// TIA Portal V19 export
FUNCTION_BLOCK "ALL_AI"   // FB2, FBD
{ S7_Optimized_Access := 'TRUE' }
// stored: MemoryReserve 100, SetENOAutomatically false
   VAR
      AI_TT01 { S7_SetPoint := 'True'} : "AI";
      TT_01 { S7_SetPoint := 'True'} : "AI";
      TT_02 { S7_SetPoint := 'True'} : "AI";
      TT_03 { S7_SetPoint := 'True'} : "AI";
      APT01 { S7_SetPoint := 'True'} : "AI";
      GPT01 { S7_SetPoint := 'True'} : "AI";
      GPT02 { S7_SetPoint := 'True'} : "AI";
      GPT03 { S7_SetPoint := 'True'} : "AI";
      GPT04 { S7_SetPoint := 'True'} : "AI";
      O201 { S7_SetPoint := 'True'} : "AI";
      LEL01 { S7_SetPoint := 'True'} : "AI";
      LEL02 { S7_SetPoint := 'True'} : "AI";
      PS01 { S7_SetPoint := 'True'} : "AI";
      RLT01 { S7_SetPoint := 'True'} : "AI";
      Weighing { S7_SetPoint := 'True'} : "AI";
   END_VAR
BEGIN

REGION Network 1: TT01
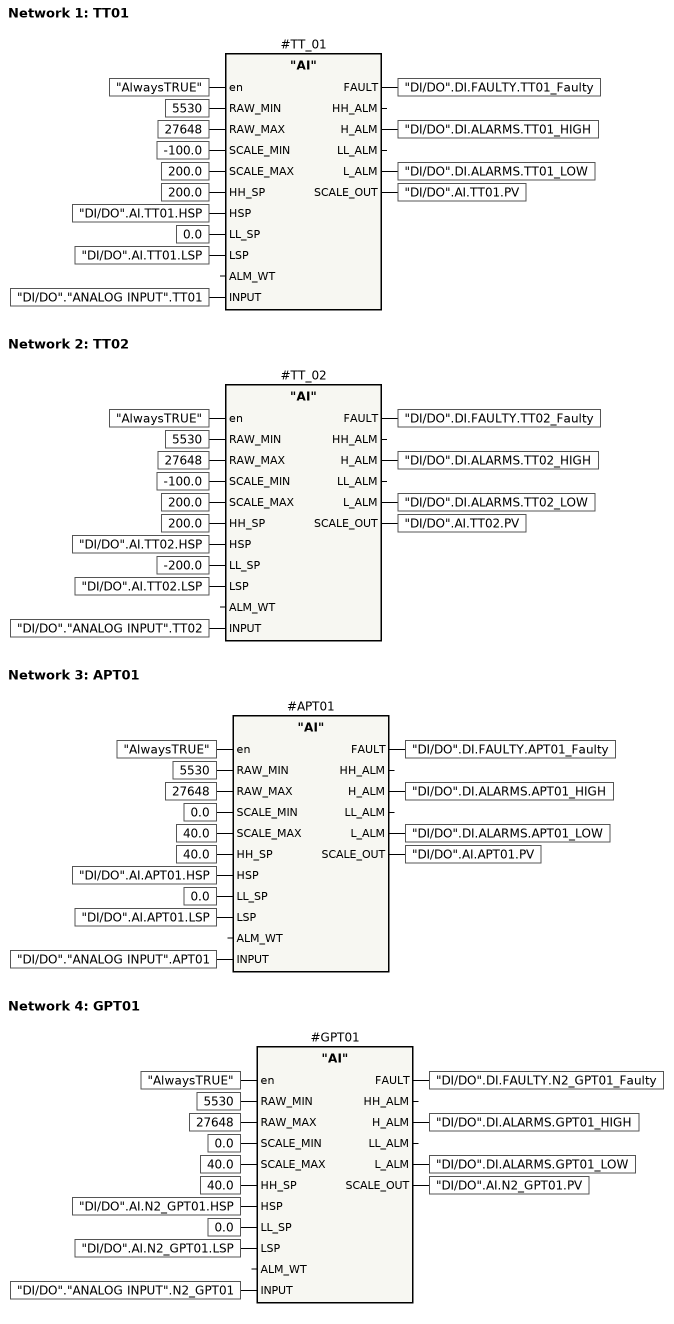
   IF "AlwaysTRUE" THEN
       #TT_01(RAW_MIN := 5530,   // "AI"
              RAW_MAX := 27648,
              SCALE_MIN := -100.0,
              SCALE_MAX := 200.0,
              HH_SP := 200.0,
              HSP := "DI/DO".AI.TT01.HSP,
              LL_SP := 0.0,
              LSP := "DI/DO".AI.TT01.LSP,
              INPUT := "DI/DO"."ANALOG INPUT".TT01,
              FAULT => "DI/DO".DI.FAULTY.TT01_Faulty,
              H_ALM => "DI/DO".DI.ALARMS.TT01_HIGH,
              L_ALM => "DI/DO".DI.ALARMS.TT01_LOW,
              SCALE_OUT => "DI/DO".AI.TT01.PV);
   END_IF;
END_REGION

REGION Network 2: TT02
   IF "AlwaysTRUE" THEN
       #TT_02(RAW_MIN := 5530,   // "AI"
              RAW_MAX := 27648,
              SCALE_MIN := -100.0,
              SCALE_MAX := 200.0,
              HH_SP := 200.0,
              HSP := "DI/DO".AI.TT02.HSP,
              LL_SP := -200.0,
              LSP := "DI/DO".AI.TT02.LSP,
              INPUT := "DI/DO"."ANALOG INPUT".TT02,
              FAULT => "DI/DO".DI.FAULTY.TT02_Faulty,
              H_ALM => "DI/DO".DI.ALARMS.TT02_HIGH,
              L_ALM => "DI/DO".DI.ALARMS.TT02_LOW,
              SCALE_OUT => "DI/DO".AI.TT02.PV);
   END_IF;
END_REGION

REGION Network 3: APT01
   IF "AlwaysTRUE" THEN
       #APT01(RAW_MIN := 5530,   // "AI"
              RAW_MAX := 27648,
              SCALE_MIN := 0.0,
              SCALE_MAX := 40.0,
              HH_SP := 40.0,
              HSP := "DI/DO".AI.APT01.HSP,
              LL_SP := 0.0,
              LSP := "DI/DO".AI.APT01.LSP,
              INPUT := "DI/DO"."ANALOG INPUT".APT01,
              FAULT => "DI/DO".DI.FAULTY.APT01_Faulty,
              H_ALM => "DI/DO".DI.ALARMS.APT01_HIGH,
              L_ALM => "DI/DO".DI.ALARMS.APT01_LOW,
              SCALE_OUT => "DI/DO".AI.APT01.PV);
   END_IF;
END_REGION

REGION Network 4: GPT01
   IF "AlwaysTRUE" THEN
       #GPT01(RAW_MIN := 5530,   // "AI"
              RAW_MAX := 27648,
              SCALE_MIN := 0.0,
              SCALE_MAX := 40.0,
              HH_SP := 40.0,
              HSP := "DI/DO".AI.N2_GPT01.HSP,
              LL_SP := 0.0,
              LSP := "DI/DO".AI.N2_GPT01.LSP,
              INPUT := "DI/DO"."ANALOG INPUT".N2_GPT01,
              FAULT => "DI/DO".DI.FAULTY.N2_GPT01_Faulty,
              H_ALM => "DI/DO".DI.ALARMS.GPT01_HIGH,
              L_ALM => "DI/DO".DI.ALARMS.GPT01_LOW,
              SCALE_OUT => "DI/DO".AI.N2_GPT01.PV);
   END_IF;
END_REGION

REGION Network 5: GPT02
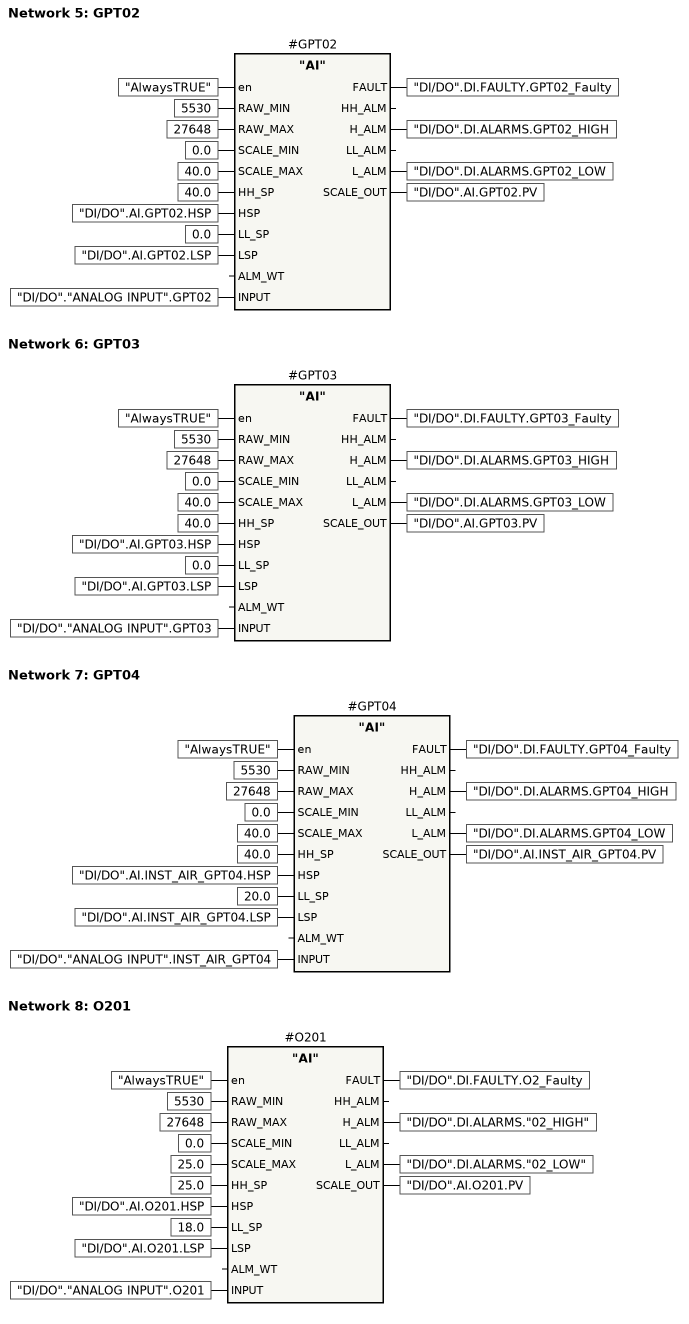
   IF "AlwaysTRUE" THEN
       #GPT02(RAW_MIN := 5530,   // "AI"
              RAW_MAX := 27648,
              SCALE_MIN := 0.0,
              SCALE_MAX := 40.0,
              HH_SP := 40.0,
              HSP := "DI/DO".AI.GPT02.HSP,
              LL_SP := 0.0,
              LSP := "DI/DO".AI.GPT02.LSP,
              INPUT := "DI/DO"."ANALOG INPUT".GPT02,
              FAULT => "DI/DO".DI.FAULTY.GPT02_Faulty,
              H_ALM => "DI/DO".DI.ALARMS.GPT02_HIGH,
              L_ALM => "DI/DO".DI.ALARMS.GPT02_LOW,
              SCALE_OUT => "DI/DO".AI.GPT02.PV);
   END_IF;
END_REGION

REGION Network 6: GPT03
   IF "AlwaysTRUE" THEN
       #GPT03(RAW_MIN := 5530,   // "AI"
              RAW_MAX := 27648,
              SCALE_MIN := 0.0,
              SCALE_MAX := 40.0,
              HH_SP := 40.0,
              HSP := "DI/DO".AI.GPT03.HSP,
              LL_SP := 0.0,
              LSP := "DI/DO".AI.GPT03.LSP,
              INPUT := "DI/DO"."ANALOG INPUT".GPT03,
              FAULT => "DI/DO".DI.FAULTY.GPT03_Faulty,
              H_ALM => "DI/DO".DI.ALARMS.GPT03_HIGH,
              L_ALM => "DI/DO".DI.ALARMS.GPT03_LOW,
              SCALE_OUT => "DI/DO".AI.GPT03.PV);
   END_IF;
END_REGION

REGION Network 7: GPT04
   IF "AlwaysTRUE" THEN
       #GPT04(RAW_MIN := 5530,   // "AI"
              RAW_MAX := 27648,
              SCALE_MIN := 0.0,
              SCALE_MAX := 40.0,
              HH_SP := 40.0,
              HSP := "DI/DO".AI.INST_AIR_GPT04.HSP,
              LL_SP := 20.0,
              LSP := "DI/DO".AI.INST_AIR_GPT04.LSP,
              INPUT := "DI/DO"."ANALOG INPUT".INST_AIR_GPT04,
              FAULT => "DI/DO".DI.FAULTY.GPT04_Faulty,
              H_ALM => "DI/DO".DI.ALARMS.GPT04_HIGH,
              L_ALM => "DI/DO".DI.ALARMS.GPT04_LOW,
              SCALE_OUT => "DI/DO".AI.INST_AIR_GPT04.PV);
   END_IF;
END_REGION

REGION Network 8: O201
   IF "AlwaysTRUE" THEN
       #O201(RAW_MIN := 5530,   // "AI"
             RAW_MAX := 27648,
             SCALE_MIN := 0.0,
             SCALE_MAX := 25.0,
             HH_SP := 25.0,
             HSP := "DI/DO".AI.O201.HSP,
             LL_SP := 18.0,
             LSP := "DI/DO".AI.O201.LSP,
             INPUT := "DI/DO"."ANALOG INPUT".O201,
             FAULT => "DI/DO".DI.FAULTY.O2_Faulty,
             H_ALM => "DI/DO".DI.ALARMS."02_HIGH",
             L_ALM => "DI/DO".DI.ALARMS."02_LOW",
             SCALE_OUT => "DI/DO".AI.O201.PV);
   END_IF;
END_REGION

REGION Network 9: LEL01
   // Configuration pending
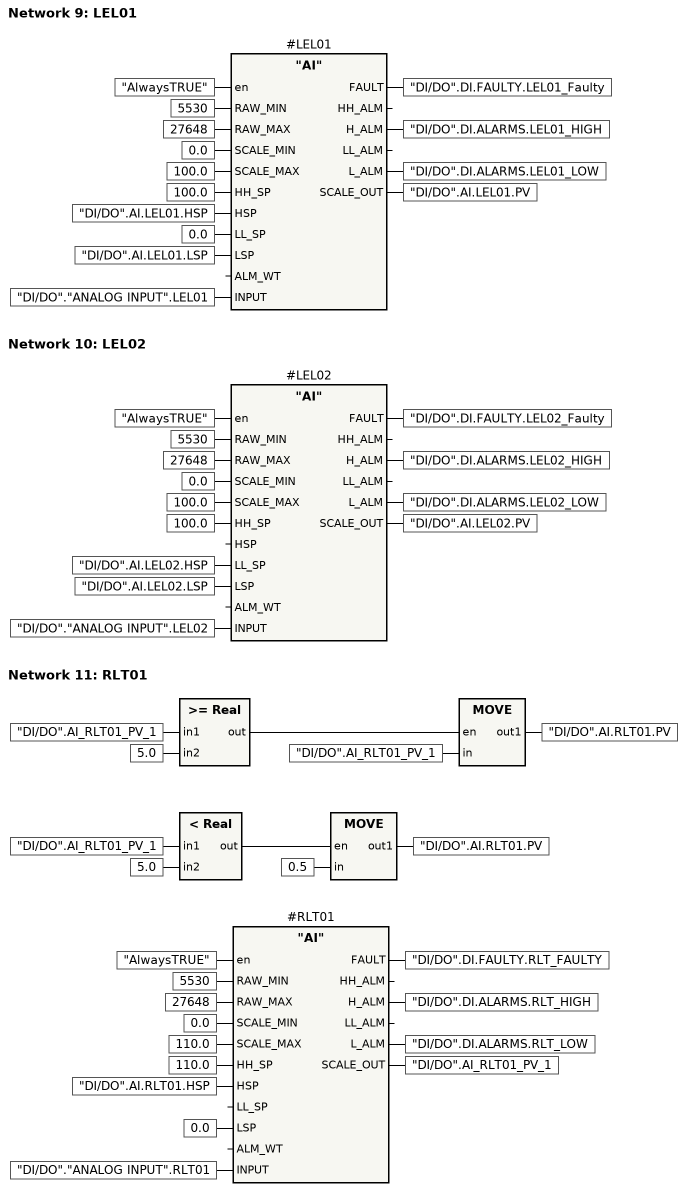
   IF "AlwaysTRUE" THEN
       #LEL01(RAW_MIN := 5530,   // "AI"
              RAW_MAX := 27648,
              SCALE_MIN := 0.0,
              SCALE_MAX := 100.0,
              HH_SP := 100.0,
              HSP := "DI/DO".AI.LEL01.HSP,
              LL_SP := 0.0,
              LSP := "DI/DO".AI.LEL01.LSP,
              INPUT := "DI/DO"."ANALOG INPUT".LEL01,
              FAULT => "DI/DO".DI.FAULTY.LEL01_Faulty,
              H_ALM => "DI/DO".DI.ALARMS.LEL01_HIGH,
              L_ALM => "DI/DO".DI.ALARMS.LEL01_LOW,
              SCALE_OUT => "DI/DO".AI.LEL01.PV);
   END_IF;
END_REGION

REGION Network 10: LEL02
   // Instrument is not installed at site
   IF "AlwaysTRUE" THEN
       #LEL02(RAW_MIN := 5530,   // "AI"
              RAW_MAX := 27648,
              SCALE_MIN := 0.0,
              SCALE_MAX := 100.0,
              HH_SP := 100.0,
              LL_SP := "DI/DO".AI.LEL02.HSP,
              LSP := "DI/DO".AI.LEL02.LSP,
              INPUT := "DI/DO"."ANALOG INPUT".LEL02,
              FAULT => "DI/DO".DI.FAULTY.LEL02_Faulty,
              H_ALM => "DI/DO".DI.ALARMS.LEL02_HIGH,
              L_ALM => "DI/DO".DI.ALARMS.LEL02_LOW,
              SCALE_OUT => "DI/DO".AI.LEL02.PV);
   END_IF;
END_REGION

REGION Network 11: RLT01
   IF "DI/DO".AI_RLT01_PV_1 >= 5.0 THEN "DI/DO".AI.RLT01.PV := "DI/DO".AI_RLT01_PV_1; END_IF;
   IF "DI/DO".AI_RLT01_PV_1 < 5.0 THEN "DI/DO".AI.RLT01.PV := 0.5; END_IF;
   IF "AlwaysTRUE" THEN
       #RLT01(RAW_MIN := 5530,   // "AI"
              RAW_MAX := 27648,
              SCALE_MIN := 0.0,
              SCALE_MAX := 110.0,
              HH_SP := 110.0,
              HSP := "DI/DO".AI.RLT01.HSP,
              LSP := 0.0,
              INPUT := "DI/DO"."ANALOG INPUT".RLT01,
              FAULT => "DI/DO".DI.FAULTY.RLT_FAULTY,
              H_ALM => "DI/DO".DI.ALARMS.RLT_HIGH,
              L_ALM => "DI/DO".DI.ALARMS.RLT_LOW,
              SCALE_OUT => "DI/DO".AI_RLT01_PV_1);
   END_IF;
END_REGION

REGION Network 12: Weighing
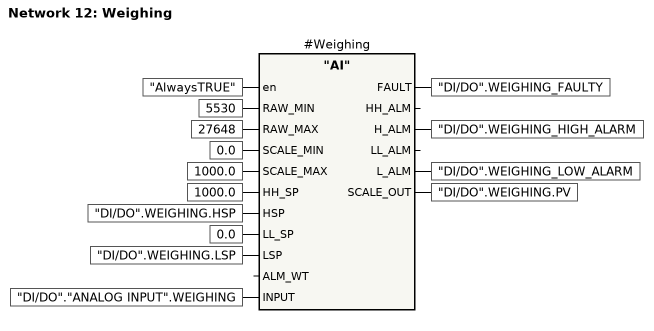
   IF "AlwaysTRUE" THEN
       #Weighing(RAW_MIN := 5530,   // "AI"
                 RAW_MAX := 27648,
                 SCALE_MIN := 0.0,
                 SCALE_MAX := 1000.0,
                 HH_SP := 1000.0,
                 HSP := "DI/DO".WEIGHING.HSP,
                 LL_SP := 0.0,
                 LSP := "DI/DO".WEIGHING.LSP,
                 INPUT := "DI/DO"."ANALOG INPUT".WEIGHING,
                 FAULT => "DI/DO".WEIGHING_FAULTY,
                 H_ALM => "DI/DO".WEIGHING_HIGH_ALARM,
                 L_ALM => "DI/DO".WEIGHING_LOW_ALARM,
                 SCALE_OUT => "DI/DO".WEIGHING.PV);
   END_IF;
END_REGION
END_FUNCTION_BLOCK
